Fanuc KAREL source: ko00060.KL

-- PROVISIONAL review KL for V770-1; original PC SHA256 11276be62a34683a9396e2350997908686790d74a30a4544c84e8b2de509e5b9
-- Incomplete behavior may be omitted. Consult companion uncertainty JSON. Do not deploy.
PROGRAM KO00060
%NOLOCKGROUP
BEGIN
  -- UNRESOLVED_PC offsets 5-12; opcodes 9D,23
  -- UNRESOLVED_PC offsets 17-69; opcodes 27,27,49,7E,AD,27,49,7E,AD,22,31,7E,4A
  -- UNRESOLVED_PC offsets 74-78; opcodes 7F
END KO00060
